// TIA Portal V20 export
Screen "IF_SIGNALS_BOOL"  1276x673
  ScreenItem "Select_InterfaceSignals" at 468,34 size 344x26  Type=HmiSymbolicIOField
  ScreenItem "Title_ScreenOverview_X390_Y2" at 390,3 size 500x30  Type=HmiTextBox
  ScreenItem "Line_Header_X0_Y64" at 0,64 size 1276x0  Type=HmiLine
  ScreenItem "Text Field_Name1" at 104,92 size 490x30  Type=HmiTextBox
  ScreenItem "Text Field_Value1" at 53,91 size 50x30  Type=HmiTextBox
  ScreenItem "Text Field_Name2" at 723,91 size 490x30  Type=HmiTextBox
  ScreenItem "Text Field_Value2" at 672,91 size 50x30  Type=HmiTextBox
  ScreenItem "EA-Feld_Free-Description_Text_Right" at 685,65 size 541x30  Type=HmiIOField
  ScreenItem "EA-Feld_Free-Description_Text_Left" at 68,66 size 541x30  Type=HmiIOField
  ScreenItem "Cycle_Time_Legend" at 1184,2 size 90x60  Type=HmiButton
  ScreenItem "permanentareaborderrectangle" at 0,0 size 0x0  Type=HmiRectangle
  ScreenItem "SymbolicName_16_Left" at 36,0 size 490x25  Type=HmiIOField
  ScreenItem "False_31" at 0,3 size 21x20  Type=HmiGraphicView
  ScreenItem "True_32" at 0,3 size 21x20  Type=HmiGraphicView
  ScreenItem "SymbolicName_15_Left" at 36,0 size 490x25  Type=HmiIOField
  ScreenItem "False_30" at 0,3 size 21x20  Type=HmiGraphicView
  ScreenItem "True_31" at 0,3 size 21x20  Type=HmiGraphicView
  ScreenItem "SymbolicName_14_Left" at 36,0 size 490x25  Type=HmiIOField
  ScreenItem "False_29" at 0,3 size 21x20  Type=HmiGraphicView
  ScreenItem "True_30" at 0,3 size 21x20  Type=HmiGraphicView
  ScreenItem "SymbolicName_13_Left" at 36,0 size 490x25  Type=HmiIOField
  ScreenItem "False_28" at 0,3 size 21x20  Type=HmiGraphicView
  ScreenItem "True_29" at 0,3 size 21x20  Type=HmiGraphicView
  ScreenItem "SymbolicName_12_Left" at 36,0 size 490x25  Type=HmiIOField
  ScreenItem "False_27" at 0,3 size 21x20  Type=HmiGraphicView
  ScreenItem "True_28" at 0,3 size 21x20  Type=HmiGraphicView
  ScreenItem "SymbolicName_11_Left" at 36,0 size 490x25  Type=HmiIOField
  ScreenItem "False_26" at 0,3 size 21x20  Type=HmiGraphicView
  ScreenItem "True_27" at 0,3 size 21x20  Type=HmiGraphicView
  ScreenItem "SymbolicName_10_Left" at 36,0 size 490x25  Type=HmiIOField
  ScreenItem "False_25" at 0,3 size 21x20  Type=HmiGraphicView
  ScreenItem "True_26" at 0,3 size 21x20  Type=HmiGraphicView
  ScreenItem "SymbolicName_9_Left" at 36,0 size 490x25  Type=HmiIOField
  ScreenItem "False_24" at 0,3 size 21x20  Type=HmiGraphicView
  ScreenItem "True_25" at 0,3 size 21x20  Type=HmiGraphicView
  ScreenItem "SymbolicName_8_Left" at 36,0 size 490x25  Type=HmiIOField
  ScreenItem "False_23" at 0,3 size 21x20  Type=HmiGraphicView
  ScreenItem "True_24" at 0,3 size 21x20  Type=HmiGraphicView
  ScreenItem "SymbolicName_7_Left" at 36,0 size 490x25  Type=HmiIOField
  ScreenItem "False_22" at 0,3 size 21x20  Type=HmiGraphicView
  ScreenItem "True_23" at 0,3 size 21x20  Type=HmiGraphicView
  ScreenItem "SymbolicName_6_Left" at 36,0 size 490x25  Type=HmiIOField
  ScreenItem "False_21" at 0,3 size 21x20  Type=HmiGraphicView
  ScreenItem "True_22" at 0,3 size 21x20  Type=HmiGraphicView
  ScreenItem "SymbolicName_5_Left" at 36,0 size 490x25  Type=HmiIOField
  ScreenItem "False_20" at 0,3 size 21x20  Type=HmiGraphicView
  ScreenItem "True_21" at 0,3 size 21x20  Type=HmiGraphicView
  ScreenItem "SymbolicName_4_Left" at 36,0 size 490x25  Type=HmiIOField
  ScreenItem "False_19" at 0,3 size 21x20  Type=HmiGraphicView
  ScreenItem "True_20" at 0,3 size 21x20  Type=HmiGraphicView
  ScreenItem "SymbolicName_3_Left" at 36,0 size 490x25  Type=HmiIOField
  ScreenItem "False_18" at 0,3 size 21x20  Type=HmiGraphicView
  ScreenItem "True_19" at 0,3 size 21x20  Type=HmiGraphicView
  ScreenItem "SymbolicName_2_Left" at 36,0 size 490x25  Type=HmiIOField
  ScreenItem "False_17" at 0,3 size 21x20  Type=HmiGraphicView
  ScreenItem "True_18" at 0,3 size 21x20  Type=HmiGraphicView
  ScreenItem "SymbolicName_1_Left" at 36,0 size 490x25  Type=HmiIOField
  ScreenItem "False_16" at 0,3 size 21x20  Type=HmiGraphicView
  ScreenItem "True_17" at 0,3 size 21x20  Type=HmiGraphicView
  ScreenItem "SymbolicName_16_Right" at 36,0 size 490x25  Type=HmiIOField
  ScreenItem "False_15" at 0,3 size 21x20  Type=HmiGraphicView
  ScreenItem "True_16" at 0,3 size 21x20  Type=HmiGraphicView
  ScreenItem "SymbolicName_15_Right" at 36,0 size 490x25  Type=HmiIOField
  ScreenItem "False_14" at 0,3 size 21x20  Type=HmiGraphicView
  ScreenItem "True_15" at 0,3 size 21x20  Type=HmiGraphicView
  ScreenItem "SymbolicName_14_Right" at 36,0 size 490x25  Type=HmiIOField
  ScreenItem "False_13" at 0,3 size 21x20  Type=HmiGraphicView
  ScreenItem "True_14" at 0,3 size 21x20  Type=HmiGraphicView
  ScreenItem "SymbolicName_13_Right" at 36,0 size 490x25  Type=HmiIOField
  ScreenItem "False_12" at 0,3 size 21x20  Type=HmiGraphicView
  ScreenItem "True_13" at 0,3 size 21x20  Type=HmiGraphicView
  ScreenItem "SymbolicName_12_Right" at 36,0 size 490x25  Type=HmiIOField
  ScreenItem "False_11" at 0,3 size 21x20  Type=HmiGraphicView
  ScreenItem "True_12" at 0,3 size 21x20  Type=HmiGraphicView
  ScreenItem "SymbolicName_11_Right" at 36,0 size 490x25  Type=HmiIOField
  ScreenItem "False_10" at 0,3 size 21x20  Type=HmiGraphicView
  ScreenItem "True_11" at 0,3 size 21x20  Type=HmiGraphicView
  ScreenItem "SymbolicName_10_Right" at 36,0 size 490x25  Type=HmiIOField
  ScreenItem "False_9" at 0,3 size 21x20  Type=HmiGraphicView
  ScreenItem "True_10" at 0,3 size 21x20  Type=HmiGraphicView
  ScreenItem "SymbolicName_9_Right" at 36,0 size 490x25  Type=HmiIOField
  ScreenItem "False_8" at 0,3 size 21x20  Type=HmiGraphicView
  ScreenItem "True_9" at 0,3 size 21x20  Type=HmiGraphicView
  ScreenItem "SymbolicName_8_Right" at 36,0 size 490x25  Type=HmiIOField
  ScreenItem "False_7" at 0,3 size 21x20  Type=HmiGraphicView
  ScreenItem "True_8" at 0,3 size 21x20  Type=HmiGraphicView
  ScreenItem "SymbolicName_7_Right" at 36,0 size 490x25  Type=HmiIOField
  ScreenItem "False_6" at 0,3 size 21x20  Type=HmiGraphicView
  ScreenItem "True_7" at 0,3 size 21x20  Type=HmiGraphicView
  ScreenItem "SymbolicName_6_Right" at 36,0 size 490x25  Type=HmiIOField
  ScreenItem "False_5" at 0,3 size 21x20  Type=HmiGraphicView
  ScreenItem "True_6" at 0,3 size 21x20  Type=HmiGraphicView
  ScreenItem "SymbolicName_5_Right" at 36,0 size 490x25  Type=HmiIOField
  ScreenItem "False_4" at 0,3 size 21x20  Type=HmiGraphicView
  ScreenItem "True_5" at 0,3 size 21x20  Type=HmiGraphicView
  ScreenItem "SymbolicName_4_Right" at 36,0 size 490x25  Type=HmiIOField
  ScreenItem "False_3" at 0,3 size 21x20  Type=HmiGraphicView
  ScreenItem "True_4" at 0,3 size 21x20  Type=HmiGraphicView
  ScreenItem "SymbolicName_3_Right" at 36,0 size 490x25  Type=HmiIOField
  ScreenItem "False_2" at 0,3 size 21x20  Type=HmiGraphicView
  ScreenItem "True_3" at 0,3 size 21x20  Type=HmiGraphicView
  ScreenItem "SymbolicName_2_Right" at 36,0 size 490x25  Type=HmiIOField
  ScreenItem "False_1" at 0,3 size 21x20  Type=HmiGraphicView
  ScreenItem "True_2" at 0,3 size 21x20  Type=HmiGraphicView
  ScreenItem "SymbolicName_1_Right" at 723,118 size 490x25  Type=HmiIOField
  ScreenItem "False_0" at 687,121 size 21x20  Type=HmiGraphicView
  ScreenItem "True_1" at 687,121 size 21x20  Type=HmiGraphicView
  ScreenItem "Button_Back" at 2,2 size 90x60  Type=HmiButton
